Fanuc KAREL source: kd00050.KL

-- PROVISIONAL review KL for V770-1; original PC SHA256 e9c7b4661df95dcbf99e0a0a2a811aed03243464d8375f6fe947203505de92ba
-- Incomplete behavior may be omitted. Consult companion uncertainty JSON. Do not deploy.
PROGRAM KD00050
%NOLOCKGROUP
VAR
  I : INTEGER
  J : INTEGER
  B : BOOLEAN
  R : REAL
  S : STRING[80]
BEGIN
  -- UNRESOLVED_PC offsets 5-19; opcodes 01,9D,2E,0A,82,0B
  -- UNRESOLVED_PC offsets 24-28; opcodes 7F
END KD00050
